// TIA Portal V20 export
DATA_BLOCK "POS3_0_Parameter_Data_Drehachse"   // DB92
{ S7_Optimized_Access := 'TRUE' }
// stored: MemoryReserve 100
   VAR
      WR_ParameterID : Word := 16#0126;
      WR_ParameterData : DWord := 16#0000_0064;
      RD_ParameterID : Word := 16#0126;
      RD_ParameterData : DWord := 16#0000_03E8;
   END_VAR
BEGIN
END_DATA_BLOCK
